FUNCTION_BLOCK TcoSingleAxis EXTENDS TcoCore.TcoComponent IMPLEMENTS ITcoSingleAxis
VAR_INPUT
	inEnable : BOOL;
    inEnablePositive : BOOL;
    inEnableNegative : BOOL;
    inCalibrationCam : BOOL;
	refAxis : REFERENCE TO TcoAxisRef;
END_VAR
VAR_IN_OUT
	inoPositions:TcoSingleAxisPositionsRootContainer;
END_VAR
VAR
	 {attribute 'hide'}
    _axisRef : REFERENCE TO TcoAxisRef;
	{attribute addProperty Name "<#Axis#>"}
	_axis :   TcoDriveSimple(THIS^);
	{attribute addProperty Name "<#Load positions Task#>"}
	_loadPositionTask :   TcoAxisExchangeDataTask(THIS^);
	{attribute addProperty Name "<#Save positions Task#>"}
	_savePositionTask :   TcoAxisExchangeDataTask(THIS^);
	{attribute addProperty Name "<#Positions#>"}
	{attribute clr [MemberByIdentity()]}
	_positions : TcoSingleAxisPositionsRootContainer(THIS^);
	{attribute addProperty Name "<#Move absolute Task#>"}
	_moveAbsoluteTask :   TcoCore.TcoTask (THIS^);
	{attribute addProperty Name "<#Move relative Task#>"}
	_moveRelativeTask :   TcoCore.TcoTask (THIS^);

	
	{attribute addProperty Name "<#Restore Task#>"}
	_restoreTask :   TcoCore.TcoTask (THIS^);
	{attribute addProperty Name "<#Status#>"}
    {attribute clr [ReadOnly()]}
    _status : TcoSingleAxisStatus;
	{attribute addProperty Name "<#Config#>"}
    _config : TcoSingleAxisConfig;
	_moveParams: TcoSingleAxisMoveParam;
	{attribute 'hide'} 
	_infoTimer :  TON;
    {attribute 'hide'} 
	_errorTimer :  TON;
END_VAR

_positions := inoPositions;

IF NOT __ISVALIDREF(refAxis)  THEN
    Messenger.Post('<#Invalid reference axis #>', TcoCore.eMessageCategory.ProgrammingError);
    RETURN;
END_IF
_axisRef REF= refAxis;


_savePositionTask();
_loadPositionTask();	

_axis(
	inEnable:=inEnable , 
	inEnablePositive:=inEnablePositive , 
	inEnableNegative:=inEnableNegative , 
	inCalibrationCam:=inCalibrationCam, 
	inoAxisRef:= _axisRef);

//*************MOVE ABSOLUTE********************
_moveAbsoluteTask.Enabled:=NOT _moveRelativeTask.Busy; 
IF _moveAbsoluteTask.Execute() THEN
	

		
	THIS^._axis.MoveAbsolute(inPosition:=_moveParams.Position,
												inVelocity:=_moveParams.Velocity,
												inAcceleration:=_moveParams.Acceleration,
												inDeceleration:=_moveParams.Deceleration,		
												inJerk:=_moveParams.Jerk);
	

		

			
	_moveAbsoluteTask.DoneWhen(THIS^._axis.MoveAbsoluteTask.Done);
	_moveAbsoluteTask.ThrowWhen(THIS^._axis.MoveAbsoluteTask.Error);	

END_IF;
//****************************************


//*************MOVE RELATIVE********************
_moveRelativeTask.Enabled:=NOT _moveAbsoluteTask.Busy; 
IF _moveRelativeTask.Execute() THEN
	
	THIS^._axis.MoveRelative(inDistance:=_moveParams.Position,
												inVelocity:=_moveParams.Velocity,
												inAcceleration:=_moveParams.Acceleration,
												inDeceleration:=_moveParams.Deceleration,		
												inJerk:=_moveParams.Jerk);
	

	_moveRelativeTask.DoneWhen(THIS^._axis.MoveRelativeTask.Done);
	_moveRelativeTask.ThrowWhen(_errorTimer.Q OR THIS^._axis.MoveRelativeTask.Error);	

END_IF;
//****************************************





//*************RESTORE********************

_restoreTask.Enabled := TRUE;
IF _restoreTask.Execute() THEN
	Restore();
END_IF
//****************************************
	
 inoPositions :=_positions;

PROPERTY Axis : REFERENCE TO TcoDriveSimple
GET
Axis REF=_axis;
END_GET
END_PROPERTY

METHOD CallTimers
VAR_INPUT
	inValue : BOOL;
END_VAR
IF  __ISVALIDREF(Config) THEN  
_infoTimer(IN := inValue, PT := THIS^.Config.InfoTime);
_errorTimer(IN := inValue, PT := THIS^.Config.ErrorTime);
END_IF;
END_METHOD

(*~
	<docu>
		<summary>
			Gets the configuration of the Axis. 					
		</summary>			
	</docu>	
~*)
PROPERTY Config : REFERENCE TO TcoSingleAxisConfig
GET
Config REF= _config;
END_GET
END_PROPERTY

PROPERTY PUBLIC LoadPositionsTask : REFERENCE TO TcoAxisExchangeDataTask
GET
LoadPositionsTask REF= _loadPositionTask;
END_GET
END_PROPERTY

METHOD MoveAbsolute : ITcoTaskStatus
VAR_INPUT
	MoveParams : TcoSingleAxisMoveParam;
END_VAR
_moveParams:=MoveParams;
MoveAbsolute:=THIS^._moveAbsoluteTask.Invoke();
END_METHOD

PROPERTY PUBLIC MoveAbsoluteTask : REFERENCE TO TcoCore.TcoTask
GET
MoveAbsoluteTask REF=_moveAbsoluteTask;
END_GET
END_PROPERTY

METHOD MoveRelative : ITcoTaskStatus
VAR_INPUT
	MoveParams : TcoSingleAxisMoveParam;
END_VAR
_moveParams:=MoveParams;
MoveRelative:=THIS^._moveRelativeTask.Invoke();
END_METHOD

PROPERTY PUBLIC MoveRelativeTask : REFERENCE TO TcoCore.TcoTask
GET
MoveRelativeTask REF=_moveRelativeTask;
END_GET
END_PROPERTY

METHOD ResetDrive : TcoCore.ITcoTaskStatus
ResetDrive:=THIS^.Axis.Reset();
END_METHOD

(*~
	<docu>
		<summary>
			Restores this instance to the Ready state. Can be called explicitly or from within one of the restore mechanisms.	
		</summary>			
	</docu>	
~*)
METHOD  Restore : ITcoRestorable
_axis.Restore();
_restoreTask.Restore();
_savePositionTask.Restore();
_loadPositionTask.Restore();
_moveAbsoluteTask.Restore();
_moveRelativeTask.Restore();
CallTimers(FALSE);
Messenger.UnPin();
END_METHOD

PROPERTY PUBLIC SavePositionsTask : REFERENCE TO TcoAxisExchangeDataTask
GET
SavePositionsTask REF= _savePositionTask;
END_GET
END_PROPERTY

METHOD PROTECTED ServiceMode
THIS^._axis.Service();
END_METHOD

METHOD SoeReset : TcoCore.ITcoTaskStatus
SoeReset:=THIS^.Axis.SoEReset();
END_METHOD

(*~
	<docu>
		<summary>
			Gets the status of the Axis system. 					
		</summary>			
	</docu>	
~*)
PROPERTY Status : REFERENCE TO TcoSingleAxisStatus
GET
Status REF= _status;
END_GET
END_PROPERTY

END_FUNCTION_BLOCK

(* stored: Version 1.1.0.1, ProductVersion 3.1.4024.12
   POU TcoSingleAxis: Id {185b24d3-f25a-4e21-b88b-2cef8570a6ca}, SpecialFunc None
   Folder Tasks: Id {8e70240b-7b2d-0f4b-36dc-8581181f84a9}
   Property Axis: Id {afff7752-8ff5-4a6a-bbec-f2ed8a50befd}
   Get Get: Id {e127fc3c-3f90-4aa4-b69d-4652a2960be6}
   Method CallTimers: Id {0a49e5e5-97c0-0f12-142a-9bf3e067c1fc}
   Property Config: Id {df1222ea-72d5-049a-39f8-23da831666e8}
   Get Get: Id {e56e9c0c-4520-0832-01b4-c85d7919c76e}
   Property LoadPositionsTask: Id {daf6c4a2-2754-03ef-30ce-d04f82ee1d2c}
   Get Get: Id {58593eb5-875f-01d6-2914-ba92ebdb8a66}
   Method MoveAbsolute: Id {e3d5c00a-e76c-4868-85c9-ff706578a857}
   Property MoveAbsoluteTask: Id {c823d07c-b5d3-018d-1f33-9a3264abca62}
   Get Get: Id {5e7f405f-d3b3-0134-0a57-ea4887c1ef97}
   Method MoveRelative: Id {27f1f345-1e04-0346-3019-bfb9b1560ada}
   Property MoveRelativeTask: Id {4784ac79-7dd3-00da-368d-7b075008258b}
   Get Get: Id {496e91ee-c0bc-029b-3484-05a455e99e60}
   Method ResetDrive: Id {0e7b0a7a-f786-06d8-3922-516d2d347d70}
   Method Restore: Id {6b84f7f5-bd0c-02a1-2804-19ef613c96e4}
   Property SavePositionsTask: Id {01670cc4-5874-0b3f-0292-2c8fa86f88c1}
   Get Get: Id {32880dc6-5d56-0f0c-039c-126a92fcd425}
   Method ServiceMode: Id {e1df90eb-bcf6-4c99-8bb6-a097504284b8}
   Method SoeReset: Id {e2ac31e5-3d50-05ab-00bc-49c90b5da0e1}
   Property Status: Id {e0852ccd-fd4f-0f31-356f-1c11062ed8c3}
   Get Get: Id {0853f10e-8dfb-0801-1cac-8d43d6440150} *)
